// Mitsubishi GX Works2 project: pivot_arm_sorter   PLC: Q03UDE

PROGRAM MAIN
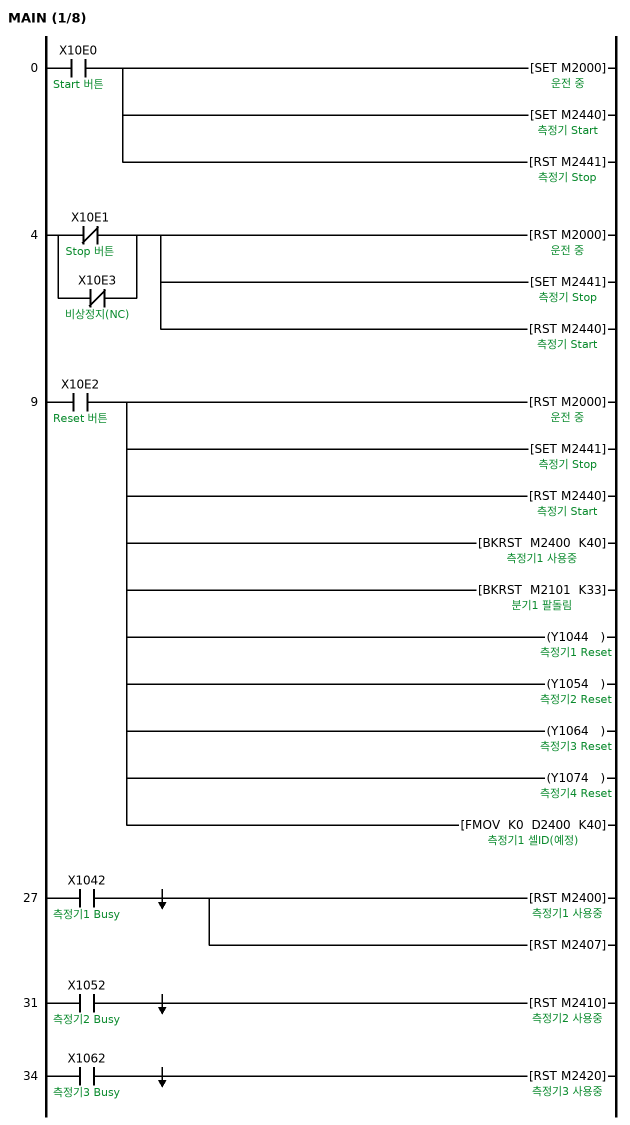
0     LD      X10E0  ; Start 버튼
      SET     M2000  ; 운전 중
      SET     M2440  ; 측정기 Start
      RST     M2441  ; 측정기 Stop
4     LDI     X10E1  ; Stop 버튼
      ORI     X10E3  ; 비상정지(NC)
      RST     M2000  ; 운전 중
      SET     M2441  ; 측정기 Stop
      RST     M2440  ; 측정기 Start
9     LD      X10E2  ; Reset 버튼
      RST     M2000  ; 운전 중
      SET     M2441  ; 측정기 Stop
      RST     M2440  ; 측정기 Start
      BKRST   M2400 K40  ; 측정기1 사용중
      BKRST   M2101 K33  ; 분기1 팔돌림
      OUT     Y1044  ; 측정기1 Reset
      OUT     Y1054  ; 측정기2 Reset
      OUT     Y1064  ; 측정기3 Reset
      OUT     Y1074  ; 측정기4 Reset
      FMOV    K0 D2400 K40  ; 측정기1 셀ID(예정)
27    LD      X1042  ; 측정기1 Busy
      MEF
      RST     M2400  ; 측정기1 사용중
      RST     M2407
31    LD      X1052  ; 측정기2 Busy
      MEF
      RST     M2410  ; 측정기2 사용중
34    LD      X1062  ; 측정기3 Busy
      MEF
      RST     M2420  ; 측정기3 사용중
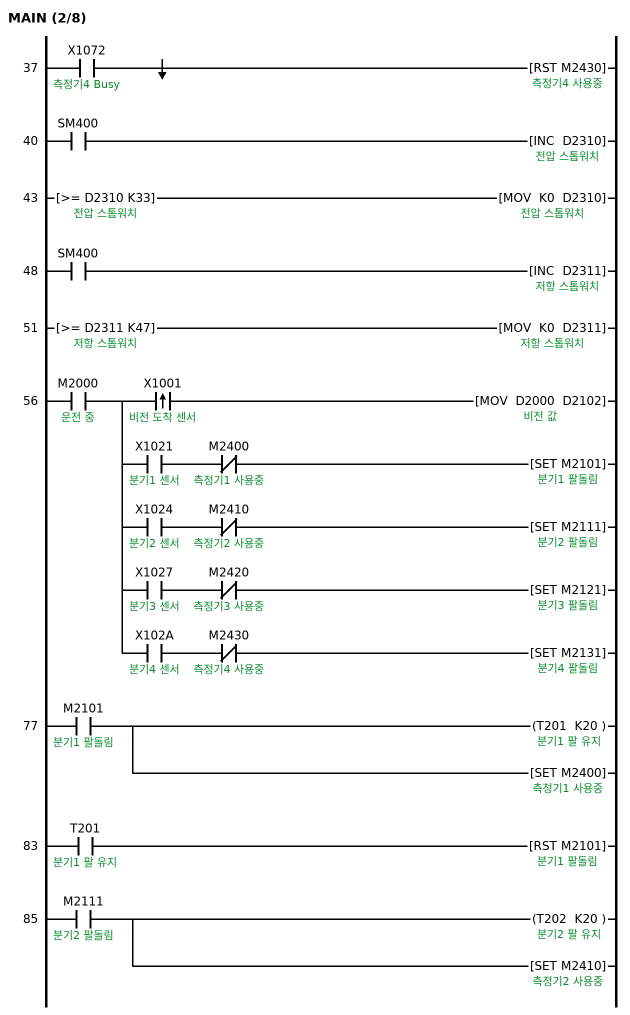
37    LD      X1072  ; 측정기4 Busy
      MEF
      RST     M2430  ; 측정기4 사용중
40    LD      SM400
      INC     D2310  ; 전압 스톱워치
43    LD>=    D2310 K33  ; 전압 스톱워치
      MOV     K0 D2310
48    LD      SM400
      INC     D2311  ; 저항 스톱워치
51    LD>=    D2311 K47  ; 저항 스톱워치
      MOV     K0 D2311
56    LD      M2000  ; 운전 중
      MPS
      ANDP    X1001  ; 비전 도착 센서
      MOV     D2000 D2102  ; 비전 값
      MRD
      AND     X1021  ; 분기1 센서
      ANI     M2400  ; 측정기1 사용중
      SET     M2101  ; 분기1 팔돌림
      MRD
      AND     X1024  ; 분기2 센서
      ANI     M2410  ; 측정기2 사용중
      SET     M2111  ; 분기2 팔돌림
      MRD
      AND     X1027  ; 분기3 센서
      ANI     M2420  ; 측정기3 사용중
      SET     M2121  ; 분기3 팔돌림
      MPP
      AND     X102A  ; 분기4 센서
      ANI     M2430  ; 측정기4 사용중
      SET     M2131  ; 분기4 팔돌림
77    LD      M2101  ; 분기1 팔돌림
      OUT     T201 K20  ; 분기1 팔 유지
      SET     M2400  ; 측정기1 사용중
83    LD      T201  ; 분기1 팔 유지
      RST     M2101  ; 분기1 팔돌림
85    LD      M2111  ; 분기2 팔돌림
      OUT     T202 K20  ; 분기2 팔 유지
      SET     M2410  ; 측정기2 사용중
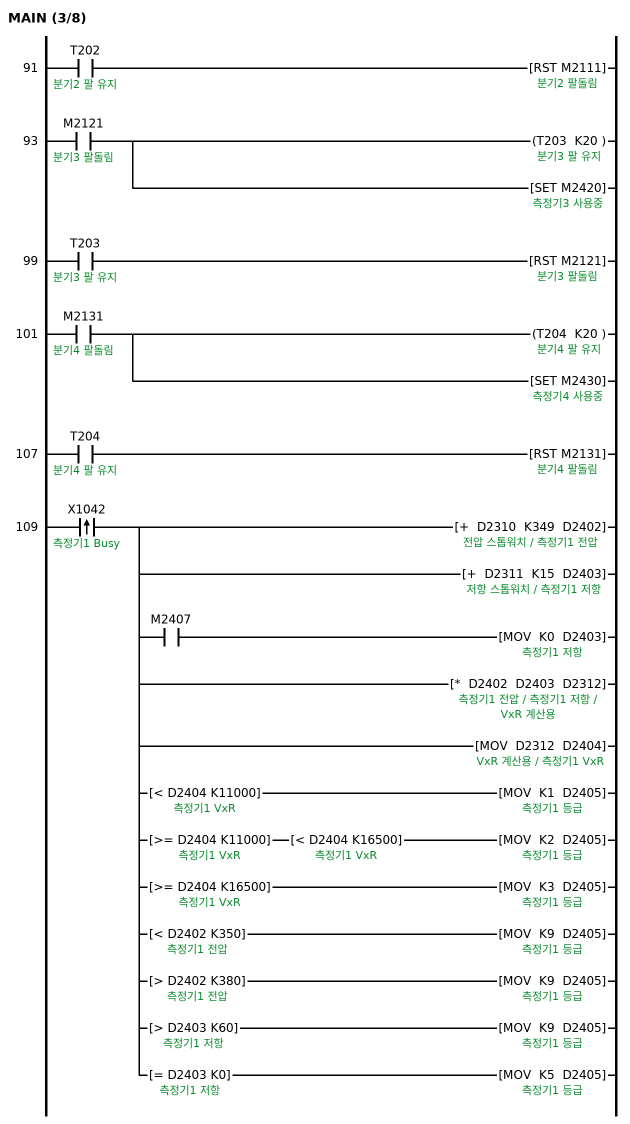
91    LD      T202  ; 분기2 팔 유지
      RST     M2111  ; 분기2 팔돌림
93    LD      M2121  ; 분기3 팔돌림
      OUT     T203 K20  ; 분기3 팔 유지
      SET     M2420  ; 측정기3 사용중
99    LD      T203  ; 분기3 팔 유지
      RST     M2121  ; 분기3 팔돌림
101   LD      M2131  ; 분기4 팔돌림
      OUT     T204 K20  ; 분기4 팔 유지
      SET     M2430  ; 측정기4 사용중
107   LD      T204  ; 분기4 팔 유지
      RST     M2131  ; 분기4 팔돌림
109   LDP     X1042  ; 측정기1 Busy
      +       D2310 K349 D2402  ; 측정기1 전압
      +       D2311 K15 D2403  ; 측정기1 저항
      MPS
      AND     M2407
      MOV     K0 D2403
      MPP
      *       D2402 D2403 D2312  ; VxR 계산용
      MOV     D2312 D2404  ; 측정기1 VxR
      MPS
      AND<    D2404 K11000  ; 측정기1 VxR
      MOV     K1 D2405  ; 측정기1 등급
      MRD
      AND>=   D2404 K11000  ; 측정기1 VxR
      AND<    D2404 K16500  ; 측정기1 VxR
      MOV     K2 D2405
      MRD
      AND>=   D2404 K16500  ; 측정기1 VxR
      MOV     K3 D2405
      MRD
      AND<    D2402 K350  ; 측정기1 전압
      MOV     K9 D2405
      MRD
      AND>    D2402 K380  ; 측정기1 전압
      MOV     K9 D2405
      MRD
      AND>    D2403 K60  ; 측정기1 저항
      MOV     K9 D2405
      MPP
      AND=    D2403 K0  ; 측정기1 저항
      MOV     K5 D2405
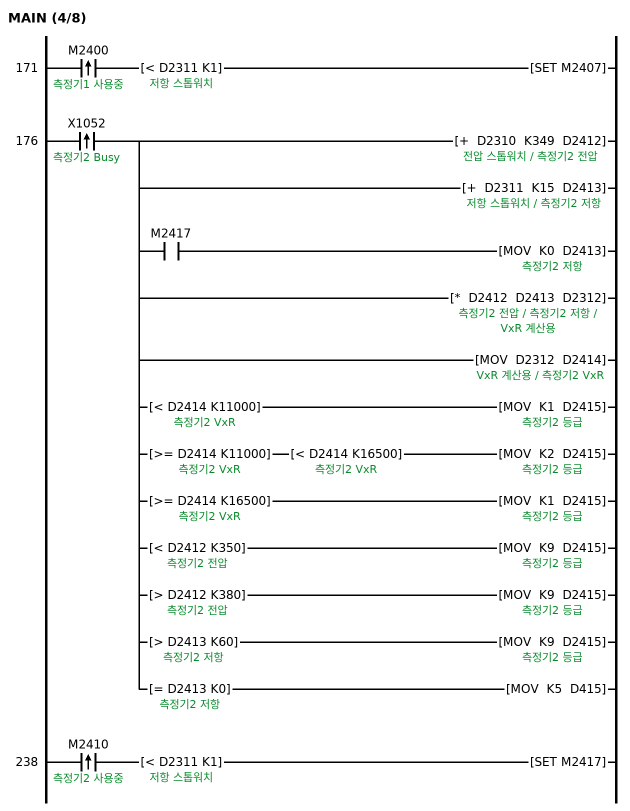
171   LDP     M2400  ; 측정기1 사용중
      AND<    D2311 K1  ; 저항 스톱워치
      SET     M2407
176   LDP     X1052  ; 측정기2 Busy
      +       D2310 K349 D2412  ; 측정기2 전압
      +       D2311 K15 D2413  ; 측정기2 저항
      MPS
      AND     M2417
      MOV     K0 D2413
      MPP
      *       D2412 D2413 D2312
      MOV     D2312 D2414  ; 측정기2 VxR
      MPS
      AND<    D2414 K11000  ; 측정기2 VxR
      MOV     K1 D2415  ; 측정기2 등급
      MRD
      AND>=   D2414 K11000  ; 측정기2 VxR
      AND<    D2414 K16500  ; 측정기2 VxR
      MOV     K2 D2415
      MRD
      AND>=   D2414 K16500  ; 측정기2 VxR
      MOV     K1 D2415
      MRD
      AND<    D2412 K350  ; 측정기2 전압
      MOV     K9 D2415
      MRD
      AND>    D2412 K380  ; 측정기2 전압
      MOV     K9 D2415
      MRD
      AND>    D2413 K60  ; 측정기2 저항
      MOV     K9 D2415
      MPP
      AND=    D2413 K0  ; 측정기2 저항
      MOV     K5 D415
238   LDP     M2410  ; 측정기2 사용중
      AND<    D2311 K1  ; 저항 스톱워치
      SET     M2417
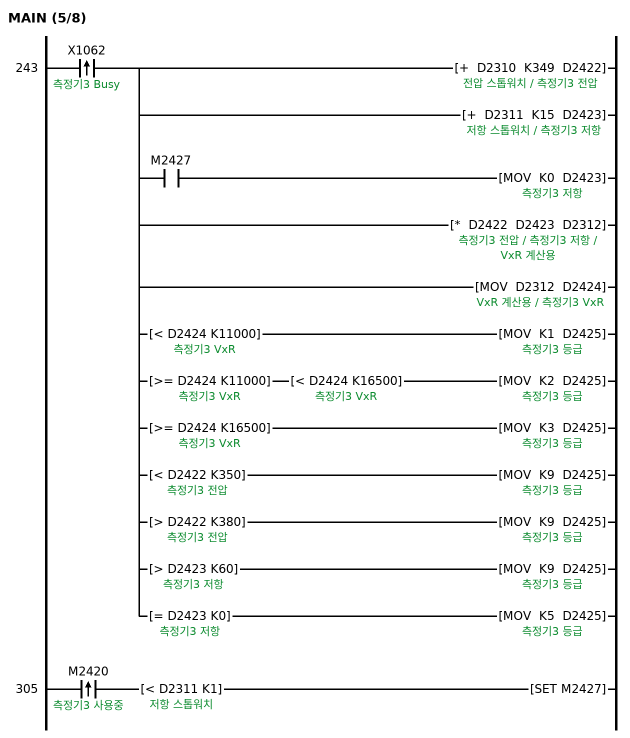
243   LDP     X1062  ; 측정기3 Busy
      +       D2310 K349 D2422  ; 측정기3 전압
      +       D2311 K15 D2423  ; 측정기3 저항
      MPS
      AND     M2427
      MOV     K0 D2423
      MPP
      *       D2422 D2423 D2312
      MOV     D2312 D2424  ; 측정기3 VxR
      MPS
      AND<    D2424 K11000  ; 측정기3 VxR
      MOV     K1 D2425  ; 측정기3 등급
      MRD
      AND>=   D2424 K11000  ; 측정기3 VxR
      AND<    D2424 K16500  ; 측정기3 VxR
      MOV     K2 D2425
      MRD
      AND>=   D2424 K16500  ; 측정기3 VxR
      MOV     K3 D2425
      MRD
      AND<    D2422 K350  ; 측정기3 전압
      MOV     K9 D2425
      MRD
      AND>    D2422 K380  ; 측정기3 전압
      MOV     K9 D2425
      MRD
      AND>    D2423 K60  ; 측정기3 저항
      MOV     K9 D2425
      MPP
      AND=    D2423 K0  ; 측정기3 저항
      MOV     K5 D2425
305   LDP     M2420  ; 측정기3 사용중
      AND<    D2311 K1  ; 저항 스톱워치
      SET     M2427
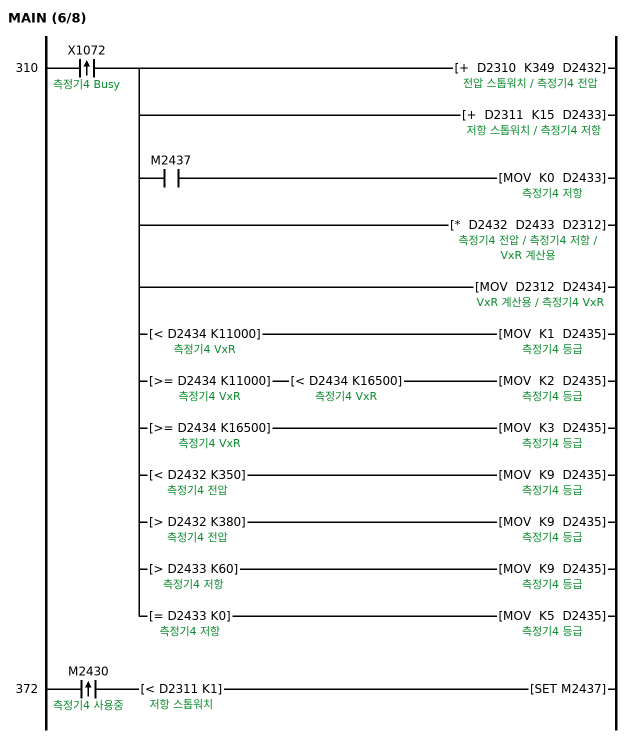
310   LDP     X1072  ; 측정기4 Busy
      +       D2310 K349 D2432  ; 측정기4 전압
      +       D2311 K15 D2433  ; 측정기4 저항
      MPS
      AND     M2437
      MOV     K0 D2433
      MPP
      *       D2432 D2433 D2312
      MOV     D2312 D2434  ; 측정기4 VxR
      MPS
      AND<    D2434 K11000  ; 측정기4 VxR
      MOV     K1 D2435  ; 측정기4 등급
      MRD
      AND>=   D2434 K11000  ; 측정기4 VxR
      AND<    D2434 K16500  ; 측정기4 VxR
      MOV     K2 D2435
      MRD
      AND>=   D2434 K16500  ; 측정기4 VxR
      MOV     K3 D2435
      MRD
      AND<    D2432 K350  ; 측정기4 전압
      MOV     K9 D2435
      MRD
      AND>    D2432 K380  ; 측정기4 전압
      MOV     K9 D2435
      MRD
      AND>    D2433 K60  ; 측정기4 저항
      MOV     K9 D2435
      MPP
      AND=    D2433 K0  ; 측정기4 저항
      MOV     K5 D2435
372   LDP     M2430  ; 측정기4 사용중
      AND<    D2311 K1  ; 저항 스톱워치
      SET     M2437
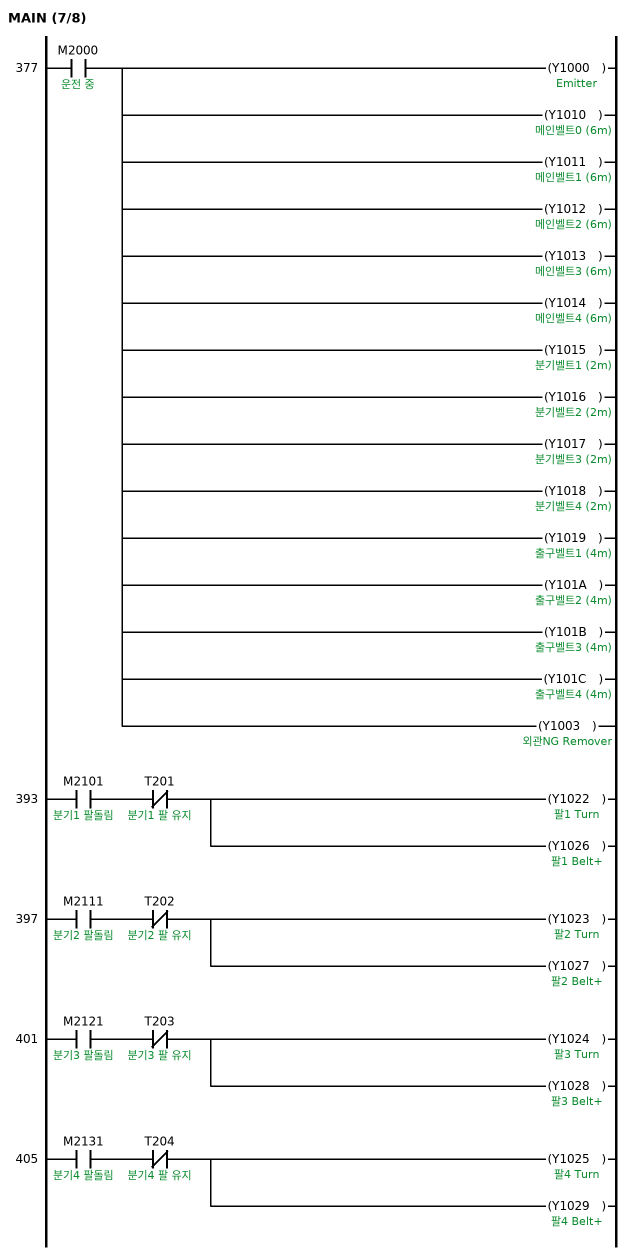
377   LD      M2000  ; 운전 중
      OUT     Y1000  ; Emitter
      OUT     Y1010  ; 메인벨트0 (6m)
      OUT     Y1011  ; 메인벨트1 (6m)
      OUT     Y1012  ; 메인벨트2 (6m)
      OUT     Y1013  ; 메인벨트3 (6m)
      OUT     Y1014  ; 메인벨트4 (6m)
      OUT     Y1015  ; 분기벨트1 (2m)
      OUT     Y1016  ; 분기벨트2 (2m)
      OUT     Y1017  ; 분기벨트3 (2m)
      OUT     Y1018  ; 분기벨트4 (2m)
      OUT     Y1019  ; 출구벨트1 (4m)
      OUT     Y101A  ; 출구벨트2 (4m)
      OUT     Y101B  ; 출구벨트3 (4m)
      OUT     Y101C  ; 출구벨트4 (4m)
      OUT     Y1003  ; 외관NG Remover
393   LD      M2101  ; 분기1 팔돌림
      ANI     T201  ; 분기1 팔 유지
      OUT     Y1022  ; 팔1 Turn
      OUT     Y1026  ; 팔1 Belt+
397   LD      M2111  ; 분기2 팔돌림
      ANI     T202  ; 분기2 팔 유지
      OUT     Y1023  ; 팔2 Turn
      OUT     Y1027  ; 팔2 Belt+
401   LD      M2121  ; 분기3 팔돌림
      ANI     T203  ; 분기3 팔 유지
      OUT     Y1024  ; 팔3 Turn
      OUT     Y1028  ; 팔3 Belt+
405   LD      M2131  ; 분기4 팔돌림
      ANI     T204  ; 분기4 팔 유지
      OUT     Y1025  ; 팔4 Turn
      OUT     Y1029  ; 팔4 Belt+
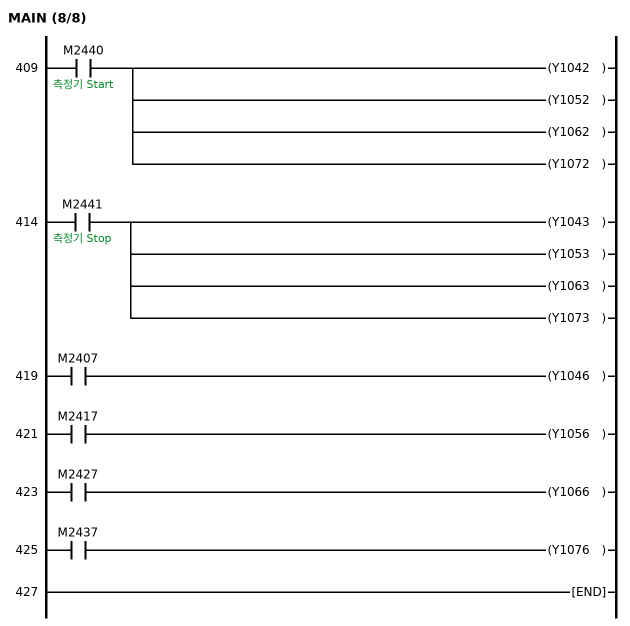
409   LD      M2440  ; 측정기 Start
      OUT     Y1042
      OUT     Y1052
      OUT     Y1062
      OUT     Y1072
414   LD      M2441  ; 측정기 Stop
      OUT     Y1043
      OUT     Y1053
      OUT     Y1063
      OUT     Y1073
419   LD      M2407
      OUT     Y1046
421   LD      M2417
      OUT     Y1056
423   LD      M2427
      OUT     Y1066
425   LD      M2437
      OUT     Y1076
427   END
END_PROGRAM

// device comments not shown above
X1000  ; 투입 센서
X1002  ; 외관NG 도착 센서
X1003  ; 외관NG 푸셔 전진끝
X1004  ; 외관NG 푸셔 복귀끝
X1020  ; 분배게이트(미사용)
X1040  ; 측정기1 입구
X1041  ; 측정기1 출구
X1043  ; 측정기1 Error
X1050  ; 측정기2 입구
X1051  ; 측정기2 출구
X1053  ; 측정기2 Error
X1060  ; 측정기3 입구
X1061  ; 측정기3 출구
X1063  ; 측정기3 Error
X1070  ; 측정기4 입구
X1071  ; 측정기4 출구
X1073  ; 측정기4 Error
Y1001  ; (예비)
Y1002  ; (예비)
Y1020  ; 분배게이트(미사용)
M2100  ; 비전 통과
M2102  ; 분기1 센서통과
M2112  ; 분기2 센서통과
M2122  ; 분기3 센서통과
M2132  ; 분기4 센서통과
M2402  ; 측정기1 측정완료
M2412  ; 측정기2 측정완료
M2422  ; 측정기3 측정완료
M2432  ; 측정기4 측정완료
D2313  ; VxR 계산용(상위)
D2401  ; 측정기1 LOT(예정)
D2410  ; 측정기2 셀ID(예정)
D2411  ; 측정기2 LOT(예정)
D2420  ; 측정기3 셀ID(예정)
D2421  ; 측정기3 LOT(예정)
D2430  ; 측정기4 셀ID(예정)
D2431  ; 측정기4 LOT(예정)
